(* IEC 61131-3 sources: rust-plc/tests/e2e-deploy/fixtures/test-project-v2, 2 files *)

(* ---- helper.st ---- *)
FUNCTION_BLOCK Accumulator
VAR
    total : INT := 0;
END_VAR
VAR_INPUT
    value : INT;
END_VAR
    total := total + value;
END_FUNCTION_BLOCK

(* ---- main.st ---- *)
(* V2: Same variable layout as V1 — compatible for online change.
   counter increments by 2 instead of 1. *)
PROGRAM Main
VAR
    counter : INT := 0;
    cycle_active : BOOL := TRUE;
END_VAR
    counter := counter + 2;
END_PROGRAM
